FUNCTION_BLOCK FB_GenericLoad IMPLEMENTS I_FeedLoad, I_JsonSource
VAR_INPUT
    stCfg : ST_GenericLoadConfig;  // this load's row of GVL_Config.aLoads
END_VAR
VAR_OUTPUT
    fAcPowerW   : LREAL;  // W at the load
    fCableLossW : LREAL;  // W lost in the load's cable, on top of fAcPowerW
END_VAR

IF stCfg.bEnabled THEN
    fAcPowerW := MAX(0.0, stCfg.fRatedPowerW);
ELSE
    fAcPowerW := 0.0;
END_IF
fCableLossW := F_CableLossW(fPowerW := fAcPowerW, fLengthFt := stCfg.fWireLengthFt, nAwg := stCfg.nWireAwg);

METHOD GetDemand : ST_LoadDemand
VAR
    stDemand : ST_LoadDemand;
END_VAR
stDemand.eKind        := E_LoadKind.Rated;
stDemand.fAcPowerW    := fAcPowerW + fCableLossW;
stDemand.fCableLossW  := fCableLossW;
stDemand.fWeight      := 0.0;
stDemand.fCableFactor := F_CableFactor(fLengthFt := stCfg.fWireLengthFt, nAwg := stCfg.nWireAwg);
stDemand.bValid       := TRUE;
GetDemand := stDemand;
END_METHOD

METHOD SetShare
VAR_INPUT
    fShareW     : LREAL;
    bShareValid : BOOL;
END_VAR
// A rated load takes no share. The method exists because I_FeedLoad requires it.
;
END_METHOD

METHOD WriteJson
VAR_INPUT
    eSection : E_JsonSection;
END_VAR
VAR_IN_OUT
    fbJson : FB_JsonSaxWriter;
END_VAR
VAR
    sFeed : STRING(20);
END_VAR
IF eSection <> E_JsonSection.Load THEN
    RETURN;
END_IF

sFeed := F_FeedIdString(nFeedId := stCfg.nFeedId);

fbJson.AddKey('id');
fbJson.AddString(stCfg.sId);
fbJson.AddKey('name');
fbJson.AddString(stCfg.sName);
fbJson.AddKey('feed');
fbJson.AddString(sFeed);
F_JsonNum(sKey := 'ratedW', fValue := stCfg.fRatedPowerW, bValid := TRUE, nDecimals := 0, fbJson := fbJson);
fbJson.AddKey('on');
fbJson.AddBool(stCfg.bEnabled);
F_JsonNum(sKey := 'cableLossW', fValue := fCableLossW, bValid := TRUE, nDecimals := 1, fbJson := fbJson);
END_METHOD

END_FUNCTION_BLOCK

(* stored: Version 1.1.0.1
   POU FB_GenericLoad: Id {81206029-0bf4-4449-9598-2df62091607f}, SpecialFunc None
   Method GetDemand: Id {ee1d4dfe-af16-4a50-a7cc-63aad0f8d55b}
   Method SetShare: Id {58371d6a-c6e3-4a2f-bbe1-7130a556f46f}
   Method WriteJson: Id {53cadb08-a563-4c86-a640-34f108fc6153} *)
